Fanuc KAREL source: kb00048.KL

-- PROVISIONAL review KL for V770-1; original PC SHA256 fd98c3bc2c5fd15229b499d32387afba8049bfebc75ac7e907d3c60f6241b0ec
-- Incomplete behavior may be omitted. Consult companion uncertainty JSON. Do not deploy.
PROGRAM KB00048
%NOLOCKGROUP
VAR
  P1 : REAL
  RESULT : REAL
BEGIN
  -- UNRESOLVED_PC offsets 5-16; opcodes 2E,23
  -- UNRESOLVED_PC offsets 21-36; opcodes 27,22,76,23
  -- UNRESOLVED_PC offsets 41-45; opcodes 7F
END KB00048
